(*
SPDX-FileCopyrightText: © 2026 Oleksandr Tiutyk <trofimich@gmail.com>
SPDX-License-Identifier: MIT
License: https://opensource.org/license/mit
*)

(*!
<summary>Validates that a generic descriptor has the configured type tag.</summary>
<description>
FB_init stores the expected tag. Validate checks exact TypeClass equality only, without dereferencing or
converting payloads; it does not validate address, size, lifetime or numeric range.
</description>
*)

{attribute 'no_explicit_call' := 'do not call this function block directly'}
FUNCTION_BLOCK GenericValueTypeValidator EXTENDS Object IMPLEMENTS IGenericValueValidator
VAR_STAT
	//! <summary>Class name shared by all instances of this function block.</summary>
	_ClassName : STRING := __POUNAME();
END_VAR
VAR
	_TypeClass : GENERIC_TYPE_CLASS;
END_VAR

{attribute 'monitoring' := 'call'}
PROPERTY ClassName : REFERENCE TO STRING
GET
ClassName REF= _ClassName;
END_GET
END_PROPERTY

(*!
<summary>Stores the exact type tag required by validation.</summary>
<description>Copies typeClass without allocating or raising exceptions. Does not inspect a value.</description>
*)
METHOD FB_init : BOOL
VAR_INPUT
	bInitRetains : BOOL; // TRUE: the retain variables are initialized (reset warm / reset cold)
	bInCopyCode : BOOL;  // TRUE: the instance will be copied to the copy code afterward (online change)
	typeClass : GENERIC_TYPE_CLASS;
END_VAR
_TypeClass := typeClass;
END_METHOD

(*!
<summary>Provides the library namespace used in diagnostics.</summary>
<description>
Borrowed read-only reference to the compiler-initialized library namespace; no ownership transfer.
</description>
*)
{attribute 'monitoring' := 'call'}
PROPERTY NamespaceName : REFERENCE TO STRING
GET
NamespaceName REF= CurrentNamespace.Name;
END_GET
END_PROPERTY

(*!
<summary>Reports the byte size of this concrete instance.</summary>
<description>
Uses XSIZEOF on the instance. Does not include separately allocated payloads or prove that an arbitrary
address is valid.
</description>
*)
{attribute 'monitoring' := 'call'}
PROPERTY SelfSize : ULINT
GET
SelfSize := XSIZEOF(THIS^);
END_GET
END_PROPERTY

(*!
<summary>Requires an exact match with the configured generic type tag.</summary>
<description>
Throws IncompatibleGenericValueTypeException on mismatch, using validatedObjectName in diagnostics. Does not
convert or inspect payload bytes, address validity or lifetime; the descriptor is borrowed and unchanged.
Descendants cannot replace exact type-tag validation; implement IGenericValueValidator separately for other
validation rules.
</description>
*)
METHOD FINAL Validate
VAR_INPUT
	validatedObjectName : WSTRING;
END_VAR
VAR_IN_OUT CONSTANT
	valueToValidate : GENERIC_VALUE;
END_VAR
IF valueToValidate.TypeClass <> _TypeClass THEN
	Exceptions.ThrowIncompatibleGenericValueType(
		sourceNamespaceName := NamespaceName,
		sourceClassName := ClassName,
		sourcePOUName := __POUNAME(),
		sourcePosition := __POSITION(),
		validatedObjectName := validatedObjectName,
		actualTypeClass := valueToValidate.TypeClass,
		expectedTypeClass := _TypeClass
	);
END_IF
END_METHOD

END_FUNCTION_BLOCK

(* stored: Version 1.1.0.1
   POU GenericValueTypeValidator: Id {a6d5904d-3010-444c-98c8-80a1917cd203}, SpecialFunc None
   Property ClassName: Id {f82f2d1b-4fc3-4718-8a54-251f7a3461ed}
   Get Get: Id {f8ee5778-fbfa-4295-aae4-9ccdc19eabec}
   Method FB_init: Id {95506783-a7ce-4b15-8e1c-b1e7f4fba622}
   Property NamespaceName: Id {9a354a72-0f79-490e-939d-4595cd41c7d6}
   Get Get: Id {81f4a78c-70ec-4b46-b623-1fc67f33b3d4}
   Property SelfSize: Id {449e46a9-6074-482b-8702-4da704e912dd}
   Get Get: Id {4b470976-567f-4fd3-acda-2171efc07a0c}
   Method Validate: Id {340dfa6e-d672-4daf-b2d9-ef30de77ce10} *)
